Yaskawa INFORM job: movjdiem.JBI

/JOB
//NAME MOVJDIEM
//POS
///NPOS 1,0,0,0,0,0
///TOOL 9
///POSTYPE PULSE
///PULSE
C00000=2100,13137,-20272,-1345,-57596,-111775
//INST
///ATTR SC,RW
///GROUP1 RB1
NOP
MOVJ C00000 VJ=10.00 PL=0
END
